(* IEC 61131-3 sources: SRCI_CLIENT_PLC/RobotLibrary/Library/POUs/Additional/MC_AbortMeasuringInput/Structures, 4 files *)

(* ---- AbortMeasuringInputOutCmd.st ---- *)
{attribute 'pack_mode' := '1'}
// -------------------------------------------------------------------------
//  SRCI Robot Library
// -------------------------------------------------------------------------
//
//  Object:      AbortMeasuringInputOutCmd
//  Author:      Thorsten Brach
//  Date:        2024-06-21
//
//  Description:
//
//
//  Copyright:
//    (C) 2024 Thorsten Brach. All rights reserved
//             Licensed under the MIT License.
//
//  Disclaimer:
//    This project is provided without any guarantee and can be used for
//    private and commercial purposes. Any use is at the user’s
//    own risk and responsibility.
//
// -------------------------------------------------------------------------
TYPE AbortMeasuringInputOutCmd :
STRUCT
END_STRUCT
END_TYPE

(* ---- AbortMeasuringInputParCmd.st ---- *)
{attribute 'pack_mode' := '1'}
// -------------------------------------------------------------------------
//  SRCI Robot Library
// -------------------------------------------------------------------------
//
//  Object:      AbortMeasuringInputParCmd
//  Author:      Thorsten Brach
//  Date:        2024-06-21
//
//  Description:
//
//
//  Copyright:
//    (C) 2024 Thorsten Brach. All rights reserved
//             Licensed under the MIT License.
//
//  Disclaimer:
//    This project is provided without any guarantee and can be used for
//    private and commercial purposes. Any use is at the user’s
//    own risk and responsibility.
//
// -------------------------------------------------------------------------
TYPE AbortMeasuringInputParCmd :
STRUCT
  /// Define an active measurement that is to be aborted.
  /// •  0: Abort all existing measurement
  /// • >0: Abort the measurement with the specific MeasuringID
  MeasuringID        : UINT;
END_STRUCT
END_TYPE

(* ---- AbortMeasuringInputRecvData.st ---- *)
{attribute 'pack_mode' := '1'}
// -------------------------------------------------------------------------
//  SRCI Robot Library
// -------------------------------------------------------------------------
//
//  Object:      AbortMeasuringInputRecvData
//  Author:      Thorsten Brach
//  Date:        2024-06-21
//
//  Description:
//
//
//  Copyright:
//    (C) 2024 Thorsten Brach. All rights reserved
//             Licensed under the MIT License.
//
//  Disclaimer:
//    This project is provided without any guarantee and can be used for
//    private and commercial purposes. Any use is at the user’s
//    own risk and responsibility.
//
// -------------------------------------------------------------------------
TYPE AbortMeasuringInputRecvData EXTENDS RspHeader :
STRUCT
END_STRUCT
END_TYPE

(* ---- AbortMeasuringInputSendData.st ---- *)
{attribute 'pack_mode' := '1'}
// -------------------------------------------------------------------------
//  SRCI Robot Library
// -------------------------------------------------------------------------
//
//  Object:      AbortMeasuringInputSendData
//  Author:      Thorsten Brach
//  Date:        2024-06-21
//
//  Description:
//
//
//  Copyright:
//    (C) 2024 Thorsten Brach. All rights reserved
//             Licensed under the MIT License.
//
//  Disclaimer:
//    This project is provided without any guarantee and can be used for
//    private and commercial purposes. Any use is at the user’s
//    own risk and responsibility.
//
// -------------------------------------------------------------------------
TYPE AbortMeasuringInputSendData EXTENDS CmdHeader:
STRUCT
  /// Define an active measurement that is to be aborted.
  /// •  0: Abort all existing measurement
  /// • >0: Abort the measurement with the specific MeasuringID
  MeasuringID        : UINT;
END_STRUCT
END_TYPE
